Staubli VAL3: refresh.pgx

public program refresh()
begin
  //功能：设置扭矩限值界面实时刷新调用
  if bLock==true
    sBtnUnLock="解锁"
  else
    sBtnUnLock="保存"
  endIf
end
